(*
SPDX-FileCopyrightText: c 2026 Oleksandr Tiutyk <trofimich@gmail.com>
SPDX-License-Identifier: MIT
License: https://opensource.org/license/mit
*)

(*!
<summary>Checks FIFO head, length and copy independence during enqueue.</summary>
<description>
Owns an inline queue and its copied entry payloads. Run from one task at a stable address.
Teardown clears surviving entries before publication, including after an aborted case.
</description>
*)

{attribute 'no_assign'}
{attribute 'no_explicit_call' := 'do not call this function block directly'}
FUNCTION_BLOCK StaticQueueEnqueueAndPeekTest EXTENDS TOF_Testing.SingleCycleTest
VAR_STAT
	{attribute 'hide'}
	_ClassName : STRING := __POUNAME();
END_VAR
VAR
	_Queue : TOF_Collections.Queue<3>(valueValidator := 0);
END_VAR

(*!
<summary>Checks FIFO head, length and copy independence during enqueue.</summary>
*)
METHOD PROTECTED ExecuteTest
VAR
	values : ARRAY [1..4] OF INT := [11, 22, 33, 44];
END_VAR
_Queue.EnqueueCopy(value := values[1]);
values[1] := 111;

Assert.ThatInt(
	actual := _Queue.Peek().AsInt(),
	message := "Changing the source must preserve the copied head"
).ToBe(expected := INT#11);

_Queue.EnqueueCopy(value := values[2]);

Assert.ThatInt(
	actual := _Queue.Peek().AsInt(),
	message := "Enqueueing the second entry must preserve the head"
).ToBe(expected := INT#11);

_Queue.EnqueueCopy(value := values[3]);

Assert.ThatInt(
	actual := _Queue.Peek().AsInt(),
	message := "Enqueueing the third entry must preserve the head"
).ToBe(expected := INT#11);

Assert.ThatBool(
	actual := _Queue.Full AND_THEN _Queue.Length = 3,
	message := "Only enqueue must advance length while peeking leaves the queue full"
).IsTrue();
END_METHOD

(*!
<summary>Restores the fixture before the runner publishes the result.</summary>
<description>
Also runs after an unexpected exception interrupts the case.
</description>
*)
METHOD PROTECTED AfterTest
_Queue.Clear();
END_METHOD

//! <summary>Borrows the concrete class name. Callers must not modify it.</summary>
{attribute 'monitoring' := 'call'}
PROPERTY ClassName : REFERENCE TO STRING
GET
ClassName REF= _ClassName;
END_GET
END_PROPERTY

//! <summary>Borrows the compiler-initialized namespace name. Callers must not modify it.</summary>
{attribute 'monitoring' := 'call'}
PROPERTY NamespaceName : REFERENCE TO STRING
GET
NamespaceName REF= CurrentNamespace.Name;
END_GET
END_PROPERTY

//! <summary>Reports the concrete instance size in bytes.</summary>
{attribute 'monitoring' := 'call'}
PROPERTY SelfSize : ULINT
GET
SelfSize := XSIZEOF(THIS^);
END_GET
END_PROPERTY

END_FUNCTION_BLOCK

(* stored: Version 1.1.0.1
   POU StaticQueueEnqueueAndPeekTest: Id {86c1a93f-8c1f-420e-bfb7-b3fc6b60d9fd}, SpecialFunc None
   Method ExecuteTest: Id {1bad0ab6-93fa-4a4e-93c0-a20f960f9ab9}
   Method AfterTest: Id {f36bd1f6-4940-474e-ad15-d7ce7234e465}
   Property ClassName: Id {49f86029-a3b5-46d7-b95b-2f223f8b23ff}
   Get Get: Id {a03cdd5f-5058-47f6-982f-749d50a20dbd}
   Property NamespaceName: Id {ddeebe28-8e85-470f-bc42-bcf9e3a99e02}
   Get Get: Id {9b39b332-9d9c-4b2a-87f1-28c383e2337b}
   Property SelfSize: Id {6ffba2b5-5ca5-4018-a64f-9c095bd209f6}
   Get Get: Id {33e510af-349b-4364-b4b8-11f13bc5abb7} *)
